(* IEC 61131-3 sources: sis-interlock-demo/tests/POUs/Suites/FB_Common_Test, 4 files *)

(* ---- DefaultCfgFailsSafe.method.decl.st ---- *)
// Умолчания ST_VotingCfg и ST_CemCfg — ошибка конфигурации (схема None, 0 причин)
METHOD PRIVATE DefaultCfgFailsSafe
VAR
    stVoteCfg : ST_VotingCfg;   // конфигурация группы по умолчанию
    stCemCfg  : ST_CemCfg;      // конфигурация матрицы по умолчанию
    wErr      : WORD;           // биты ошибок матрицы
END_VAR

(* ---- DefaultStsFailSafe.method.decl.st ---- *)
// Умолчания состояний: ST_VoteResult и ST_VotingSts — срабатывание без схемы; свежий FB_Voting —
// xTrip = TRUE, свежий FB_CauseEffect — xTripped = TRUE и все выходы FALSE (до первого вызова)
METHOD PRIVATE DefaultStsFailSafe
VAR
    stRes  : ST_VoteResult;    // результат по умолчанию
    stSts  : ST_VotingSts;     // состояние группы по умолчанию
    fbVote : FB_Voting;        // не вызывался
    fbCem  : FB_CauseEffect;   // не вызывался
    uiJ    : UINT;             // индекс следствия
    xAnyOn : BOOL;             // хотя бы один выход под напряжением
END_VAR

(* ---- DefaultStsFailSafe.method.impl.st ---- *)
coUnit.TEST('Common_DefaultSts_FailSafe');
AssertTrue(Condition := stRes.xTrip, Message := 'ST_VoteResult default: trip');
AssertEquals_INT(Expected := TO_INT(E_VoteArch.None), Actual := TO_INT(stRes.eArchEff),
    Message := 'ST_VoteResult default: arch None');
AssertTrue(Condition := stSts.xTrip, Message := 'ST_VotingSts default: trip');
AssertTrue(Condition := fbVote.xTrip, Message := 'FB_Voting before first call: trip');
AssertTrue(Condition := fbCem.xTripped, Message := 'FB_CauseEffect before first call: tripped');
xAnyOn := FALSE;
FOR uiJ := 1 TO GVL_Const.SIS_EFFECTS_MAX DO
    xAnyOn := xAnyOn OR fbCem.axEffectOut[uiJ];
END_FOR
AssertFalse(Condition := xAnyOn, Message := 'FB_CauseEffect before first call: all outputs de-energized');
coUnit.TEST_FINISHED();

(* ---- SizeLimitsMasksFitWord.method.decl.st ---- *)
// Маски причин и следствий — WORD: SIS_CAUSES_MAX и SIS_EFFECTS_MAX не больше 16; каналов 3; журнал 64
METHOD PRIVATE SizeLimitsMasksFitWord
VAR
    wMask : WORD;   // пример маски
END_VAR
